TYPE stSwitchState :
STRUCT
    // Logical state
    CurrentState        : eSwitchStateType;         // Current processed state
    PreviousState       : eSwitchStateType;         // Previous state
    StateChanged        : BOOL;                // State change flag
    
    // Counters
    PressCount          : USINT := 0;            // Number of clicks in sequence
    TotalPresses        : UDINT := 0;          // Total number of clicks

END_STRUCT
END_TYPE

(* stored: Version 1.1.0.1
   DUT stSwitchState: Id {95f89ab6-dc0c-4e63-95ce-633bc21eb204} *)
